(* IEC 61131-3 sources: plc-process-lib/tests/POUs/Suites/FB_Alarm_Test, 48 files *)

(* ---- AckAfterReturnGoesNormal.method.decl.st ---- *)
// Квитирование вернувшейся тревоги: RtnUnack → Normal, тревога уходит из списка.
METHOD PRIVATE AckAfterReturnGoesNormal
VAR
    fbTime : FB_FakeTime;    // подменное время
    fbAlm  : FB_Alarm;       // ФБ под тестом
    stCfg  : ST_AlarmCfg;    // параметры по умолчанию
    xRet   : BOOL;           // ответ метода
END_VAR

(* ---- AckAndClearSameCallTwoEventsInOrder.method.decl.st ---- *)
// Квитирование и уход условия в одном вызове: два перехода по порядку шагов тела — Acked
// (ActiveUnack → ActiveAck), затем Cleared (ActiveAck → Normal); udiSeq + 2.
METHOD PRIVATE AckAndClearSameCallTwoEventsInOrder
VAR
    fbTime : FB_FakeTime;    // подменное время
    fbAlm  : FB_Alarm;       // ФБ под тестом
    stCfg  : ST_AlarmCfg;    // параметры по умолчанию
    fbSink : FB_TestSink;    // приёмник событий
    stEv   : ST_AlarmEvent;  // прочитанное событие
END_VAR

(* ---- AckInNormalReturnsFalse.method.decl.st ---- *)
// Ack без эффекта: в Normal и ActiveAck метод возвращает FALSE и переходов не даёт.
METHOD PRIVATE AckInNormalReturnsFalse
VAR
    fbTime : FB_FakeTime;    // подменное время
    fbAlm  : FB_Alarm;       // ФБ под тестом
    stCfg  : ST_AlarmCfg;    // параметры по умолчанию
    xRet   : BOOL;           // ответ Ack
END_VAR

(* ---- AckWhileActiveGoesActiveAck.method.decl.st ---- *)
// Квитирование активной тревоги: Ack() возвращает TRUE и только ставит запрос; ближайший вызов
// тела переводит ActiveUnack → ActiveAck (тревога остаётся в списке, неквитированности нет).
METHOD PRIVATE AckWhileActiveGoesActiveAck
VAR
    fbTime : FB_FakeTime;    // подменное время
    fbAlm  : FB_Alarm;       // ФБ под тестом
    stCfg  : ST_AlarmCfg;    // параметры по умолчанию
    xRet   : BOOL;           // ответ метода
END_VAR

(* ---- AckWithoutEffectNotKeptForLater.method.decl.st ---- *)
// Квитирование без эффекта не запоминается: Ack в Normal и в Shelved выполняется ближайшим вызовом
// тела и снимается. Следующее появление тревоги (в том числе повторное оповещение после снятия
// shelve) остаётся ActiveUnack и в следующих вызовах — «заранее квитировать» тревогу нельзя
// (ISA-18.2: оператор должен увидеть каждое новое появление)
METHOD PRIVATE AckWithoutEffectNotKeptForLater
VAR
    fbTime : FB_FakeTime;    // подменное время
    fbAlm  : FB_Alarm;       // ФБ под тестом
    stCfg  : ST_AlarmCfg;    // параметры по умолчанию
END_VAR

(* ---- ActivateGoesActiveUnack.method.decl.st ---- *)
// Условие появилось (без задержек): Normal → ActiveUnack; xActive, xUnacked, xInList взведены,
// udiSeq = 1, ltLastChange — время перехода.
METHOD PRIVATE ActivateGoesActiveUnack
VAR
    fbTime : FB_FakeTime;    // подменное время, старт 1 ч
    fbAlm  : FB_Alarm;       // ФБ под тестом
    stCfg  : ST_AlarmCfg;    // Medium, без задержек, shelve до 8 ч
END_VAR

(* ---- ActiveAckReturnGoesNormal.method.decl.st ---- *)
// Квитированная активная тревога, условие ушло: ActiveAck → Normal (причина Cleared).
METHOD PRIVATE ActiveAckReturnGoesNormal
VAR
    fbTime : FB_FakeTime;    // подменное время
    fbAlm  : FB_Alarm;       // ФБ под тестом
    stCfg  : ST_AlarmCfg;    // параметры по умолчанию
    fbSink : FB_TestSink;    // приёмник событий
    stEv   : ST_AlarmEvent;  // последнее событие
END_VAR

(* ---- ActiveWhileShelvedFollowsCondition.method.decl.st ---- *)
// xActive показывает условие после задержек независимо от наложенного состояния: при shelve
// условие уходит и возвращается — xActive следует за ним, состояние Shelved не меняется.
METHOD PRIVATE ActiveWhileShelvedFollowsCondition
VAR
    fbTime : FB_FakeTime;    // подменное время
    fbAlm  : FB_Alarm;       // ФБ под тестом
    stCfg  : ST_AlarmCfg;    // параметры по умолчанию
    itfAlm : I_Alarm;        // тот же ФБ через интерфейс
END_VAR

(* ---- InterfacePropertiesMatchOutputs.method.decl.st ---- *)
// Свойства I_Alarm совпадают с выходами ФБ: Id, State, AlarmPriority, Active, Unacked, Seq.
METHOD PRIVATE InterfacePropertiesMatchOutputs
VAR
    fbTime : FB_FakeTime;    // подменное время
    fbAlm  : FB_Alarm;       // ФБ под тестом
    stCfg  : ST_AlarmCfg;    // приоритет Low
    itfAlm : I_Alarm;        // тот же ФБ через интерфейс
END_VAR

(* ---- NonFiniteValueEventValueFinite.method.decl.st ---- *)
// Значение процесса NaN в момент перехода (PV из Modbus): rValue события конечно — 0.0 (R6: приёмник журнала и SQL
// не получают NaN); конечное значение передаётся как есть.
METHOD PRIVATE NonFiniteValueEventValueFinite
VAR
    fbTime : FB_FakeTime;    // подменное время
    fbAlm  : FB_Alarm;       // ФБ под тестом
    stCfg  : ST_AlarmCfg;    // умолчания (Medium)
    fbSink : FB_TestSink;    // приёмник событий
    stEv1  : ST_AlarmEvent;  // событие при NaN
    stEv2  : ST_AlarmEvent;  // событие при конечном значении
    uBits  : U_RealBits;     // NaN по битам
END_VAR

(* ---- NoTimeSourceFallsBackToSystemTime.method.decl.st ---- *)
// Без источника (itfTime = 0) FB_Alarm берёт встроенный FB_SystemTime: тревога без задержки
// появляется сразу, отметка перехода больше 0; задержка 1 ч за время теста не истекает.
METHOD PRIVATE NoTimeSourceFallsBackToSystemTime
VAR
    fbAlm  : FB_Alarm;       // без задержки
    fbAlm2 : FB_Alarm;       // задержка появления 1 ч
    stCfg  : ST_AlarmCfg;    // параметры по умолчанию
    iStep  : INT;            // шаг цикла
END_VAR

(* ---- NoTimeSourceFallsBackToSystemTime.method.impl.st ---- *)
coUnit.TEST('Alarm_NoTimeSource_FallsBackToSystemTime');

fbAlm(xIn := TRUE, stCfg := stCfg);
AssertTrue(Condition := fbAlm.eState = E_AlarmState.ActiveUnack, Message := 'activated with system time');
AssertTrue(Condition := fbAlm.ltLastChange > LTIME#0S, Message := 'system time stamp above zero');
stCfg.tOnDelay := T#1H;
FOR iStep := 1 TO 100 DO
    fbAlm2(xIn := TRUE, stCfg := stCfg);
END_FOR
AssertTrue(Condition := fbAlm2.eState = E_AlarmState.Normal, Message := 'on-delay of 1 h does not expire');

coUnit.TEST_FINISHED();

(* ---- OffDelayHoldsActive.method.decl.st ---- *)
// Задержка снятия 2 с: после ухода условия тревога остаётся ActiveUnack до 1,9 с и переходит в
// RtnUnack ровно в 2,0 с.
METHOD PRIVATE OffDelayHoldsActive
VAR
    fbTime : FB_FakeTime;    // подменное время
    fbAlm  : FB_Alarm;       // ФБ под тестом
    stCfg  : ST_AlarmCfg;    // tOffDelay = 2 с
    iStep  : INT;            // шаг цикла
END_VAR

(* ---- OffDelayHoldsActive.method.impl.st ---- *)
coUnit.TEST('Alarm_OffDelay_HoldsActive');

stCfg.tOffDelay := T#2S;
fbAlm(xIn := TRUE, stCfg := stCfg, itfTime := fbTime);                                // ActiveUnack сразу
AssertTrue(Condition := fbAlm.eState = E_AlarmState.ActiveUnack, Message := 'no on-delay: active at once');
fbTime.Advance(tStep := T#1S);
fbAlm(xIn := FALSE, stCfg := stCfg, itfTime := fbTime);                               // t1: условие ушло
FOR iStep := 1 TO 19 DO                                                               // до t1 + 1,9 с
    fbTime.Advance(tStep := T#100MS);
    fbAlm(xIn := FALSE, stCfg := stCfg, itfTime := fbTime);
END_FOR
AssertTrue(Condition := fbAlm.eState = E_AlarmState.ActiveUnack, Message := 'still active at t1 + 1.9 s');
AssertTrue(Condition := fbAlm.xActive, Message := 'xActive held by the off-delay');
fbTime.Advance(tStep := T#100MS);
fbAlm(xIn := FALSE, stCfg := stCfg, itfTime := fbTime);                               // t1 + 2,0 с
AssertTrue(Condition := fbAlm.eState = E_AlarmState.RtnUnack, Message := 'RtnUnack exactly at t1 + 2.0 s');

coUnit.TEST_FINISHED();

(* ---- OnDelayShortConditionNoAlarm.method.decl.st ---- *)
// Задержка появления 3 с: условие 2,9 с тревоги не даёт; устойчивое условие — ActiveUnack ровно
// через 3,0 с (на шаге 2,9 с ещё Normal).
METHOD PRIVATE OnDelayShortConditionNoAlarm
VAR
    fbTime  : FB_FakeTime;   // подменное время
    fbAlm   : FB_Alarm;      // ФБ под тестом
    stCfg   : ST_AlarmCfg;   // tOnDelay = 3 с
    xEver   : BOOL;          // тревога хоть раз ушла из Normal
    iStep   : INT;           // шаг цикла
END_VAR

(* ---- OnDelayShortConditionNoAlarm.method.impl.st ---- *)
coUnit.TEST('Alarm_OnDelay_ShortCondition_NoAlarm');

stCfg.tOnDelay := T#3S;
fbAlm(xIn := TRUE, stCfg := stCfg, itfTime := fbTime);                                // t0: условие
FOR iStep := 1 TO 29 DO                                                               // до t0 + 2,9 с
    fbTime.Advance(tStep := T#100MS);
    fbAlm(xIn := TRUE, stCfg := stCfg, itfTime := fbTime);
    xEver := xEver OR fbAlm.eState <> E_AlarmState.Normal;
END_FOR
FOR iStep := 1 TO 20 DO                                                               // условие ушло
    fbTime.Advance(tStep := T#100MS);
    fbAlm(xIn := FALSE, stCfg := stCfg, itfTime := fbTime);
    xEver := xEver OR fbAlm.eState <> E_AlarmState.Normal;
END_FOR
AssertFalse(Condition := xEver, Message := 'condition of 2.9 s with tOnDelay 3 s raises no alarm');
AssertEquals_UDINT(Expected := 0, Actual := fbAlm.udiSeq, Message := 'no transitions');

fbAlm(xIn := TRUE, stCfg := stCfg, itfTime := fbTime);                                // t1: условие
FOR iStep := 1 TO 29 DO
    fbTime.Advance(tStep := T#100MS);
    fbAlm(xIn := TRUE, stCfg := stCfg, itfTime := fbTime);
END_FOR
AssertTrue(Condition := fbAlm.eState = E_AlarmState.Normal, Message := 'no alarm at t1 + 2.9 s');
fbTime.Advance(tStep := T#100MS);
fbAlm(xIn := TRUE, stCfg := stCfg, itfTime := fbTime);                                // t1 + 3,0 с
AssertTrue(Condition := fbAlm.eState = E_AlarmState.ActiveUnack, Message := 'alarm exactly at t1 + 3.0 s');

coUnit.TEST_FINISHED();

(* ---- OosEntryClearsUnackReannunciatesOnExit.method.decl.st ---- *)
// Вход в OutOfService из ActiveUnack снимает неквитированность; при выходе с активным условием
// тревога снова ActiveUnack, без условия — Normal.
METHOD PRIVATE OosEntryClearsUnackReannunciatesOnExit
VAR
    fbTime : FB_FakeTime;    // подменное время
    fbAlm  : FB_Alarm;       // с активным условием
    fbAlm2 : FB_Alarm;       // условие уходит во время OutOfService
    stCfg  : ST_AlarmCfg;    // параметры по умолчанию
END_VAR

(* ---- OosOffWithSuppressActiveGoesSuppressed.method.decl.st ---- *)
// Выход из OutOfService при действующем подавлении — SuppressedByDesign (причина OosOff), а не
// базовое состояние.
METHOD PRIVATE OosOffWithSuppressActiveGoesSuppressed
VAR
    fbTime : FB_FakeTime;    // подменное время
    fbAlm  : FB_Alarm;       // ФБ под тестом
    stCfg  : ST_AlarmCfg;    // параметры по умолчанию
    fbSink : FB_TestSink;    // приёмник событий
    stEv   : ST_AlarmEvent;  // последнее событие
END_VAR

(* ---- OutOfServiceOverridesShelve.method.decl.st ---- *)
// OutOfService старше shelve: отложенная тревога уходит в OutOfService, срок shelve продолжает
// идти (xShelved = TRUE); Shelve в OutOfService не принимается. Выход из OutOfService до конца
// срока — снова Shelved с остатком 40 мин; срок, истёкший в OutOfService, — при выходе базовое
// состояние (условие активно — ActiveUnack).
METHOD PRIVATE OutOfServiceOverridesShelve
VAR
    fbTime : FB_FakeTime;    // подменное время
    fbAlm  : FB_Alarm;       // ФБ под тестом
    stCfg  : ST_AlarmCfg;    // параметры по умолчанию
    fbSink : FB_TestSink;    // приёмник событий
    stEv   : ST_AlarmEvent;  // последнее событие
    xRet   : BOOL;           // ответ Shelve
END_VAR

(* ---- PriorityChangeWhileActiveNoEvent.method.decl.st ---- *)
// Смена приоритета активной тревоги (Medium → High) действует сразу и события не порождает.
METHOD PRIVATE PriorityChangeWhileActiveNoEvent
VAR
    fbTime : FB_FakeTime;    // подменное время
    fbAlm  : FB_Alarm;       // ФБ под тестом
    stCfg  : ST_AlarmCfg;    // Medium, затем High
    itfAlm : I_Alarm;        // тот же ФБ через интерфейс
END_VAR

(* ---- PriorityNoneCancelsShelve.method.decl.st ---- *)
// Выключение тревоги (приоритет None) снимает действующий shelve: Normal с событием Disabled (ALM-1),
// xShelved = FALSE, остаток 0. После включения при активном условии — Activated (ActiveUnack), а не Shelved:
// shelve выключенной тревоги не «доживает» до её включения. Контракт 10.2, F-21 (б)
METHOD PRIVATE PriorityNoneCancelsShelve
VAR
    fbTime : FB_FakeTime;    // подменное время
    fbAlm  : FB_Alarm;       // ФБ под тестом
    stCfg  : ST_AlarmCfg;    // Medium, затем None, затем снова Medium
    fbSink : FB_TestSink;    // приёмник событий
    stEv   : ST_AlarmEvent;  // последнее событие
    udiSeq : UDINT;          // udiSeq до выключения
END_VAR

(* ---- PriorityNoneNeverActivates.method.decl.st ---- *)
// Приоритет None выключает тревогу: при активном условии 10 вызовов — Normal, все выходы FALSE,
// udiSeq = 0, событий нет; Shelve и Ack — FALSE.
METHOD PRIVATE PriorityNoneNeverActivates
VAR
    fbTime : FB_FakeTime;    // подменное время
    fbAlm  : FB_Alarm;       // ФБ под тестом
    stCfg  : ST_AlarmCfg;    // приоритет None
    fbSink : FB_TestSink;    // приёмник событий
    xEver  : BOOL;           // хоть раз взведён какой-либо выход
    xRet   : BOOL;           // ответы методов
    iStep  : INT;            // шаг цикла
END_VAR

(* ---- PriorityNoneNeverActivates.method.impl.st ---- *)
coUnit.TEST('Alarm_PriorityNone_NeverActivates');

stCfg.ePriority := E_AlarmPriority.None;
GVL_Lib.itfAlarmSink := fbSink;
FOR iStep := 1 TO 10 DO
    fbAlm(xIn := TRUE, stCfg := stCfg, itfTime := fbTime);
    xEver := xEver OR fbAlm.xActive OR fbAlm.xUnacked OR fbAlm.xInList OR fbAlm.xShelved
             OR fbAlm.eState <> E_AlarmState.Normal;
    fbTime.Advance(tStep := T#1S);
END_FOR
GVL_Lib.itfAlarmSink := 0;
xRet := fbAlm.Shelve(tDuration := T#0S) OR fbAlm.Ack();
AssertFalse(Condition := xEver, Message := 'disabled alarm: Normal, all outputs FALSE');
AssertEquals_UDINT(Expected := 0, Actual := fbAlm.udiSeq, Message := 'udiSeq unchanged');
AssertEquals_UINT(Expected := 0, Actual := fbSink.Count, Message := 'no events');
AssertFalse(Condition := xRet, Message := 'Shelve and Ack return FALSE');

coUnit.TEST_FINISHED();

(* ---- PriorityNoneToMediumActiveConditionActivates.method.decl.st ---- *)
// Включение выключенной тревоги при активном условии: приоритет None → Medium даёт Activated в
// том же вызове (без задержки); с tOnDelay 1 с — через 1 с после включения.
METHOD PRIVATE PriorityNoneToMediumActiveConditionActivates
VAR
    fbTime : FB_FakeTime;    // подменное время
    fbAlm  : FB_Alarm;       // без задержки
    fbAlm2 : FB_Alarm;       // с задержкой появления
    stCfg  : ST_AlarmCfg;    // приоритет None, затем Medium
    iStep  : INT;            // шаг цикла
END_VAR

(* ---- PriorityNoneToMediumActiveConditionActivates.method.impl.st ---- *)
coUnit.TEST('Alarm_PriorityNoneToMedium_ActiveCondition_Activates');

stCfg.ePriority := E_AlarmPriority.None;
FOR iStep := 1 TO 5 DO
    fbAlm(xIn := TRUE, stCfg := stCfg, itfTime := fbTime);
    fbTime.Advance(tStep := T#1S);
END_FOR
stCfg.ePriority := E_AlarmPriority.Medium;
fbAlm(xIn := TRUE, stCfg := stCfg, itfTime := fbTime);
AssertTrue(Condition := fbAlm.eState = E_AlarmState.ActiveUnack,
           Message := 'enabled with active condition -> Activated');
AssertEquals_UDINT(Expected := 1, Actual := fbAlm.udiSeq, Message := 'one transition');

stCfg.ePriority := E_AlarmPriority.None;
stCfg.tOnDelay := T#1S;
FOR iStep := 1 TO 5 DO
    fbAlm2(xIn := TRUE, stCfg := stCfg, itfTime := fbTime);
    fbTime.Advance(tStep := T#1S);
END_FOR
stCfg.ePriority := E_AlarmPriority.Medium;
fbAlm2(xIn := TRUE, stCfg := stCfg, itfTime := fbTime);                               // t1: включена
AssertTrue(Condition := fbAlm2.eState = E_AlarmState.Normal, Message := 'on-delay starts at enabling');
fbTime.Advance(tStep := T#1S);
fbAlm2(xIn := TRUE, stCfg := stCfg, itfTime := fbTime);                               // t1 + 1 с
AssertTrue(Condition := fbAlm2.eState = E_AlarmState.ActiveUnack, Message := 'activated 1 s after enabling');

coUnit.TEST_FINISHED();

(* ---- PriorityNoneWhileActiveEmitsClosingEvent.method.decl.st ---- *)
// Тревога ActiveUnack, приоритет переключили на None (ALM-1): переход в Normal с событием Disabled (старое состояние
// ActiveUnack, новое Normal, udiSeq + 1) — журнал и сводка по событиям закрывают тревогу. Дальше выключенная
// тревога событий не даёт.
METHOD PRIVATE PriorityNoneWhileActiveEmitsClosingEvent
VAR
    fbTime : FB_FakeTime;    // подменное время
    fbAlm  : FB_Alarm;       // ФБ под тестом
    stCfg  : ST_AlarmCfg;    // Medium, затем None
    fbSink : FB_TestSink;    // приёмник событий
    stEv   : ST_AlarmEvent;  // последнее событие
    udiSeq : UDINT;          // udiSeq до выключения
    uiCnt  : UINT;           // событий после выключения
END_VAR

(* ---- PriorityOutOfEnumTreatedAsMedium.method.decl.st ---- *)
// Приоритет вне перечисления (9 — мусор persistent-памяти) не выключает тревогу: она работает как
// Medium, свойство и событие показывают Medium.
METHOD PRIVATE PriorityOutOfEnumTreatedAsMedium
VAR
    fbTime : FB_FakeTime;    // подменное время
    fbAlm  : FB_Alarm;       // ФБ под тестом
    stCfg  : ST_AlarmCfg;    // приоритет 9
    uBad   : U_TestEnumInt;  // число вне перечисления
    fbSink : FB_TestSink;    // приёмник событий
    stEv   : ST_AlarmEvent;  // последнее событие
    itfAlm : I_Alarm;        // тот же ФБ через интерфейс
END_VAR

(* ---- PriorityReenabledOnDelayCountsFromEnabling.method.decl.st ---- *)
// Задержка появления после выключения и включения тревоги отсчитывается заново, от включения:
// тревога с tOnDelay 2 с была активна и квитирована, на 5 с выключена (приоритет None) при
// активном условии; после включения — Normal 1,9 с и ActiveUnack ровно через 2 с, а не сразу по
// старому состоянию задержки. F-21 (б)
METHOD PRIVATE PriorityReenabledOnDelayCountsFromEnabling
VAR
    fbTime : FB_FakeTime;    // подменное время
    fbAlm  : FB_Alarm;       // ФБ под тестом
    stCfg  : ST_AlarmCfg;    // tOnDelay 2 с
    iStep  : INT;            // шаг цикла
END_VAR

(* ---- PriorityReenabledOnDelayCountsFromEnabling.method.impl.st ---- *)
coUnit.TEST('Alarm_PriorityReenabled_OnDelayCountsFromEnabling');

stCfg.tOnDelay := T#2S;
fbAlm(xIn := TRUE, stCfg := stCfg, itfTime := fbTime);
fbTime.Advance(tStep := T#2S);
fbAlm(xIn := TRUE, stCfg := stCfg, itfTime := fbTime);                                // ActiveUnack через 2 с
fbAlm.Ack();
fbAlm(xIn := TRUE, stCfg := stCfg, itfTime := fbTime);                                // ActiveAck
AssertTrue(Condition := fbAlm.eState = E_AlarmState.ActiveAck, Message := 'precondition: ActiveAck');
stCfg.ePriority := E_AlarmPriority.None;
FOR iStep := 1 TO 5 DO
    fbTime.Advance(tStep := T#1S);
    fbAlm(xIn := TRUE, stCfg := stCfg, itfTime := fbTime);                            // выключена, условие есть
END_FOR
stCfg.ePriority := E_AlarmPriority.Medium;
fbAlm(xIn := TRUE, stCfg := stCfg, itfTime := fbTime);                                // t1: включена
FOR iStep := 1 TO 19 DO
    fbTime.Advance(tStep := T#100MS);
    fbAlm(xIn := TRUE, stCfg := stCfg, itfTime := fbTime);
END_FOR
AssertTrue(Condition := fbAlm.eState = E_AlarmState.Normal, Message := 'Normal until t1 + 1.9 s');
AssertFalse(Condition := fbAlm.xActive, Message := 'condition not active before the on-delay');
fbTime.Advance(tStep := T#100MS);
fbAlm(xIn := TRUE, stCfg := stCfg, itfTime := fbTime);                                // t1 + 2,0 с
AssertTrue(Condition := fbAlm.eState = E_AlarmState.ActiveUnack, Message := 'ActiveUnack exactly at t1 + 2 s');

coUnit.TEST_FINISHED();

(* ---- ReactivateFromRtnUnackGoesActiveUnack.method.decl.st ---- *)
// Условие вернулось до квитирования: RtnUnack → ActiveUnack (причина Activated).
METHOD PRIVATE ReactivateFromRtnUnackGoesActiveUnack
VAR
    fbTime : FB_FakeTime;    // подменное время
    fbAlm  : FB_Alarm;       // ФБ под тестом
    stCfg  : ST_AlarmCfg;    // параметры по умолчанию
    fbSink : FB_TestSink;    // приёмник событий
    stEv   : ST_AlarmEvent;  // последнее событие
END_VAR

(* ---- ReshelveRestartsTimer.method.decl.st ---- *)
// Повторный Shelve во время shelve отсчитывает срок заново: через 40 мин после первого — снова 1 ч.
METHOD PRIVATE ReshelveRestartsTimer
VAR
    fbTime : FB_FakeTime;    // подменное время
    fbAlm  : FB_Alarm;       // ФБ под тестом
    stCfg  : ST_AlarmCfg;    // параметры по умолчанию
    xRet   : BOOL;           // ответ Shelve
END_VAR

(* ---- ReturnWithoutAckGoesRtnUnack.method.decl.st ---- *)
// Условие ушло до квитирования: ActiveUnack → RtnUnack; тревога остаётся неквитированной и в списке.
METHOD PRIVATE ReturnWithoutAckGoesRtnUnack
VAR
    fbTime : FB_FakeTime;    // подменное время
    fbAlm  : FB_Alarm;       // ФБ под тестом
    stCfg  : ST_AlarmCfg;    // параметры по умолчанию
END_VAR

(* ---- SeqIncrementsOnEachTransition.method.decl.st ---- *)
// udiSeq (и свойство Seq) растёт на 1 на каждом переходе: Activated, Acked, Shelved, Unshelved,
// Cleared, Acked — 6; вызовы без перехода счётчик не меняют.
METHOD PRIVATE SeqIncrementsOnEachTransition
VAR
    fbTime : FB_FakeTime;    // подменное время
    fbAlm  : FB_Alarm;       // ФБ под тестом
    stCfg  : ST_AlarmCfg;    // параметры по умолчанию
    itfAlm : I_Alarm;        // тот же ФБ через интерфейс
END_VAR

(* ---- ShelveDurationAboveMaxClippedToMax.method.decl.st ---- *)
// Срок shelve больше tShelveMax (2 ч при максимуме 1 ч) обрезается до максимума; меньший срок
// (30 мин) берётся как есть.
METHOD PRIVATE ShelveDurationAboveMaxClippedToMax
VAR
    fbTime : FB_FakeTime;    // подменное время
    fbAlm  : FB_Alarm;       // ФБ под тестом
    stCfg  : ST_AlarmCfg;    // tShelveMax = 1 ч
    xRet   : BOOL;           // ответ Shelve
END_VAR

(* ---- ShelveExpiresDuringSuppressReleaseGoesToBase.method.decl.st ---- *)
// Срок shelve истёк во время подавления: состояние остаётся SuppressedByDesign, xShelved снят;
// снятие подавления при активном условии — ActiveUnack.
METHOD PRIVATE ShelveExpiresDuringSuppressReleaseGoesToBase
VAR
    fbTime : FB_FakeTime;    // подменное время
    fbAlm  : FB_Alarm;       // ФБ под тестом
    stCfg  : ST_AlarmCfg;    // tShelveMax = 1 ч
END_VAR

(* ---- ShelveMaxZeroShelveRejected.method.decl.st ---- *)
// tShelveMax = T#0S запрещает shelve: Shelve() возвращает FALSE, тревога остаётся ActiveUnack.
// Выключенная тревога (приоритет None) shelve тоже не принимает.
METHOD PRIVATE ShelveMaxZeroShelveRejected
VAR
    fbTime : FB_FakeTime;    // подменное время
    fbAlm  : FB_Alarm;       // ФБ под тестом
    stCfg  : ST_AlarmCfg;    // tShelveMax = 0
    xRet   : BOOL;           // ответ Shelve
END_VAR

(* ---- ShelveRemainCountsDown.method.decl.st ---- *)
// Остаток shelve убывает со временем: shelve 1 ч, через 15 мин — 45 мин, через 59 мин 59 с — 1 с.
METHOD PRIVATE ShelveRemainCountsDown
VAR
    fbTime : FB_FakeTime;    // подменное время
    fbAlm  : FB_Alarm;       // ФБ под тестом
    stCfg  : ST_AlarmCfg;    // параметры по умолчанию
END_VAR

(* ---- ShelveRequestThenOosRejected.method.decl.st ---- *)
// Запрос Shelve принят методом (тревога ещё не в OutOfService), но в ближайшем вызове тела поднялся
// xOutOfService: тело запрос отклоняет — shelve не начинается, после выхода из OutOfService тревога
// не Shelved, а базовое состояние (условие активно — ActiveUnack). F-21 (в), контракт 10.1
METHOD PRIVATE ShelveRequestThenOosRejected
VAR
    fbTime : FB_FakeTime;    // подменное время
    fbAlm  : FB_Alarm;       // ФБ под тестом
    stCfg  : ST_AlarmCfg;    // параметры по умолчанию (tShelveMax 8 ч)
    xRet   : BOOL;           // ответ Shelve
END_VAR

(* ---- ShelveTimeoutUnshelvesAndReannunciates.method.decl.st ---- *)
// Shelve квитированной активной тревоги на tShelveMax = 8 ч (T#0S в запросе): Shelved, остаток 8 ч,
// тревога не в списке. По истечении срока при активном условии — снова ActiveUnack (повторное
// оповещение, причина ShelveExpired); в 7 ч 50 мин ещё Shelved. Шаг времени 10 мин.
METHOD PRIVATE ShelveTimeoutUnshelvesAndReannunciates
VAR
    fbTime : FB_FakeTime;    // подменное время
    fbAlm  : FB_Alarm;       // ФБ под тестом
    stCfg  : ST_AlarmCfg;    // tShelveMax = 8 ч (по умолчанию)
    fbSink : FB_TestSink;    // приёмник событий
    stEv   : ST_AlarmEvent;  // последнее событие
    xRet   : BOOL;           // ответ Shelve
    iStep  : INT;            // шаг цикла
END_VAR

(* ---- ShelveTimeoutUnshelvesAndReannunciates.method.impl.st ---- *)
coUnit.TEST('Alarm_Shelve_TimeoutUnshelvesAndReannunciates');

GVL_Lib.itfAlarmSink := fbSink;
fbAlm(xIn := TRUE, stCfg := stCfg, itfTime := fbTime);                                // ActiveUnack
fbAlm.Ack();
fbAlm(xIn := TRUE, stCfg := stCfg, itfTime := fbTime);                                // ActiveAck
xRet := fbAlm.Shelve(tDuration := T#0S);
fbAlm(xIn := TRUE, stCfg := stCfg, itfTime := fbTime);                                // t0: Shelved
AssertTrue(Condition := xRet, Message := 'shelve accepted');
AssertTrue(Condition := fbAlm.eState = E_AlarmState.Shelved, Message := 'ActiveAck -> Shelved');
AssertTrue(Condition := fbAlm.xShelved, Message := 'xShelved set');
AssertEquals_TIME(Expected := T#8H, Actual := fbAlm.tShelveRemain, Message := 'T#0S means tShelveMax = 8 h');
AssertFalse(Condition := fbAlm.xInList, Message := 'shelved alarm is not in the list');
FOR iStep := 1 TO 47 DO                                                               // до t0 + 7 ч 50 мин
    fbTime.Advance(tStep := T#10M);
    fbAlm(xIn := TRUE, stCfg := stCfg, itfTime := fbTime);
END_FOR
AssertTrue(Condition := fbAlm.eState = E_AlarmState.Shelved, Message := 'still shelved at 7 h 50 min');
AssertEquals_TIME(Expected := T#10M, Actual := fbAlm.tShelveRemain, Message := '10 min left');
fbTime.Advance(tStep := T#10M);
fbAlm(xIn := TRUE, stCfg := stCfg, itfTime := fbTime);                                // t0 + 8 ч
GVL_Lib.itfAlarmSink := 0;
AssertTrue(Condition := fbAlm.eState = E_AlarmState.ActiveUnack, Message := 'reannunciated as ActiveUnack after 8 h');
AssertFalse(Condition := fbAlm.xShelved, Message := 'shelve ended');
AssertEquals_TIME(Expected := T#0S, Actual := fbAlm.tShelveRemain, Message := 'no shelve time left');
stEv := fbSink.Last;
AssertTrue(Condition := stEv.eReason = E_AlarmEventReason.ShelveExpired, Message := 'event reason ShelveExpired');
AssertTrue(Condition := stEv.eOldState = E_AlarmState.Shelved, Message := 'event old state Shelved');

coUnit.TEST_FINISHED();

(* ---- ShelveWhileSuppressedShelvedAfterRelease.method.decl.st ---- *)
// Shelve во время подавления принимается (не OutOfService): состояние остаётся SuppressedByDesign,
// xShelved = TRUE, событий нет; снятие подавления — Shelved (причина Unsuppressed).
METHOD PRIVATE ShelveWhileSuppressedShelvedAfterRelease
VAR
    fbTime : FB_FakeTime;    // подменное время
    fbAlm  : FB_Alarm;       // ФБ под тестом
    stCfg  : ST_AlarmCfg;    // параметры по умолчанию
    fbSink : FB_TestSink;    // приёмник событий
    stEv   : ST_AlarmEvent;  // последнее событие
    xRet   : BOOL;           // ответ Shelve
END_VAR

(* ---- SuppressByDesignNoAnnunciation.method.decl.st ---- *)
// Подавление по условию: при xSuppress активная тревога — SuppressedByDesign, не в списке, не
// требует квитирования (Ack — FALSE), xActive показывает условие. Снятие подавления при активном
// условии — ActiveUnack (причина Unsuppressed): оператор видит тревогу заново.
METHOD PRIVATE SuppressByDesignNoAnnunciation
VAR
    fbTime : FB_FakeTime;    // подменное время
    fbAlm  : FB_Alarm;       // ФБ под тестом
    stCfg  : ST_AlarmCfg;    // параметры по умолчанию
    fbSink : FB_TestSink;    // приёмник событий
    stEv   : ST_AlarmEvent;  // последнее событие
    xRet   : BOOL;           // ответ Ack
    iStep  : INT;            // шаг цикла
END_VAR

(* ---- SuppressByDesignNoAnnunciation.method.impl.st ---- *)
coUnit.TEST('Alarm_SuppressByDesign_NoAnnunciation');

GVL_Lib.itfAlarmSink := fbSink;
FOR iStep := 1 TO 10 DO
    fbAlm(xIn := TRUE, xSuppress := TRUE, stCfg := stCfg, itfTime := fbTime);
    fbTime.Advance(tStep := T#1S);
END_FOR
xRet := fbAlm.Ack();
AssertTrue(Condition := fbAlm.eState = E_AlarmState.SuppressedByDesign, Message := 'suppressed by design');
AssertFalse(Condition := fbAlm.xInList, Message := 'not in the alarm list');
AssertFalse(Condition := fbAlm.xUnacked, Message := 'no acknowledge needed');
AssertFalse(Condition := xRet, Message := 'Ack has no effect while suppressed');
AssertTrue(Condition := fbAlm.xActive, Message := 'xActive shows the condition');
AssertEquals_UDINT(Expected := 1, Actual := fbAlm.udiSeq, Message := 'one transition (Normal -> SuppressedByDesign)');
fbAlm(xIn := TRUE, xSuppress := FALSE, stCfg := stCfg, itfTime := fbTime);
GVL_Lib.itfAlarmSink := 0;
AssertTrue(Condition := fbAlm.eState = E_AlarmState.ActiveUnack,
           Message := 'release with active condition -> ActiveUnack');
stEv := fbSink.Last;
AssertTrue(Condition := stEv.eReason = E_AlarmEventReason.Unsuppressed, Message := 'event reason Unsuppressed');

coUnit.TEST_FINISHED();

(* ---- SuppressClearsUnackReleaseWithoutConditionGoesNormal.method.decl.st ---- *)
// Вход в подавление сбрасывает неквитированность (ActiveUnack → SuppressedByDesign); условие ушло
// во время подавления — снятие подавления даёт Normal, а не RtnUnack.
METHOD PRIVATE SuppressClearsUnackReleaseWithoutConditionGoesNormal
VAR
    fbTime : FB_FakeTime;    // подменное время
    fbAlm  : FB_Alarm;       // ФБ под тестом
    stCfg  : ST_AlarmCfg;    // параметры по умолчанию
END_VAR

(* ---- TimeBackwardsShelveRemainNotExtended.method.decl.st ---- *)
// «Время назад» во время shelve (SetNow на 2 ч раньше): остаток не растёт сверх срока (1 ч), shelve
// заканчивается через 1 ч от нового времени.
METHOD PRIVATE TimeBackwardsShelveRemainNotExtended
VAR
    fbTime : FB_FakeTime;    // подменное время
    fbAlm  : FB_Alarm;       // ФБ под тестом
    stCfg  : ST_AlarmCfg;    // параметры по умолчанию
END_VAR

(* ---- TransitionSendsEventToSink.method.decl.st ---- *)
// Каждый переход отправляет событие в GVL_Lib.itfAlarmSink: номер, приоритет, старое и новое
// состояние, причина, отметка времени и значение процесса.
METHOD PRIVATE TransitionSendsEventToSink
VAR
    fbTime : FB_FakeTime;    // подменное время
    fbAlm  : FB_Alarm;       // ФБ под тестом
    stCfg  : ST_AlarmCfg;    // приоритет High
    fbSink : FB_TestSink;    // приёмник событий
    stEv   : ST_AlarmEvent;  // прочитанное событие
    ltAct  : LTIME;          // время появления
END_VAR

(* ---- UnshelveConditionClearedGoesNormal.method.decl.st ---- *)
// Условие ушло, пока тревога отложена: состояние Shelved, xActive = FALSE. Unshelve переводит в
// Normal (причина Unshelved), без повторного оповещения.
METHOD PRIVATE UnshelveConditionClearedGoesNormal
VAR
    fbTime : FB_FakeTime;    // подменное время
    fbAlm  : FB_Alarm;       // ФБ под тестом
    stCfg  : ST_AlarmCfg;    // параметры по умолчанию
    fbSink : FB_TestSink;    // приёмник событий
    stEv   : ST_AlarmEvent;  // последнее событие
    xRet   : BOOL;           // ответ Unshelve
END_VAR

(* ---- UnshelveReturnsTrueOnlyWhenShelved.method.decl.st ---- *)
// Unshelve возвращает TRUE, только пока shelve действует; без shelve запрос ни на что не влияет.
METHOD PRIVATE UnshelveReturnsTrueOnlyWhenShelved
VAR
    fbTime : FB_FakeTime;    // подменное время
    fbAlm  : FB_Alarm;       // ФБ под тестом
    stCfg  : ST_AlarmCfg;    // параметры по умолчанию
    xRet   : BOOL;           // ответ Unshelve
END_VAR
